Fanuc KAREL source: kt00370.KL

-- PROVISIONAL review KL for V1013-1; original PC SHA256 a1e9b71cb020b3ca6ddeca2696baac55ad39fcea7299688c6874a80156288182
-- Incomplete behavior may be omitted. Consult companion uncertainty JSON. Do not deploy.
PROGRAM KT00370
%NOLOCKGROUP
VAR
  R1 : REAL
  R2 : REAL
  OUT : BOOLEAN
BEGIN
  -- UNRESOLVED_PC offsets 5-16; opcodes 2E,23
  -- UNRESOLVED_PC offsets 21-32; opcodes 2E,23
  -- UNRESOLVED_PC offsets 37-48; opcodes 2E,23
  -- UNRESOLVED_PC offsets 53-64; opcodes 2E,23
  -- UNRESOLVED_PC offsets 69-88; opcodes 21,21,70,23
  -- UNRESOLVED_PC offsets 93-97; opcodes 7F
END KT00370
